Staubli VAL3: utList.dtx

public utAppearance Appearance
  [0]
    string sBackgroundColour
    string sColour
    bool bVisibility
public utBorder Border
  [0]
    string sBorderColour
    string sBorderStyle
    string sBorderWidth
public utCommon Common
  [0]
    bool bDisabled
    string sValue
    string sID
    string sOption{}
    string sItem
    string sPage
public utText Text
  [0]
    string sFontFamily
    string sFontStyle
    num nFontSize
